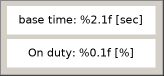
VISUALIZATION vis_FB_DutyCycle_Master  // 164x76
VAR_IN_OUT
	fBaseTime	: REAL;
	fOn_Duty	: REAL;		
END_VAR
    Rectangle (0,0 164x76)
    Textfield (6,5 150x30), "base time: %2.1f [sec]", text variable: fBaseTime
        OnMouseClick: write the text variable via Edit, min 0, max 60
    Textfield (6,38 150x30), "On duty: %0.1f [%]", text variable: fOn_Duty
        OnMouseClick: write the text variable via Edit, min 0, max 100
END_VISUALIZATION

// ---- 01 Instance/04 Recipe/Vis_Recipe_Tab.TcVIS
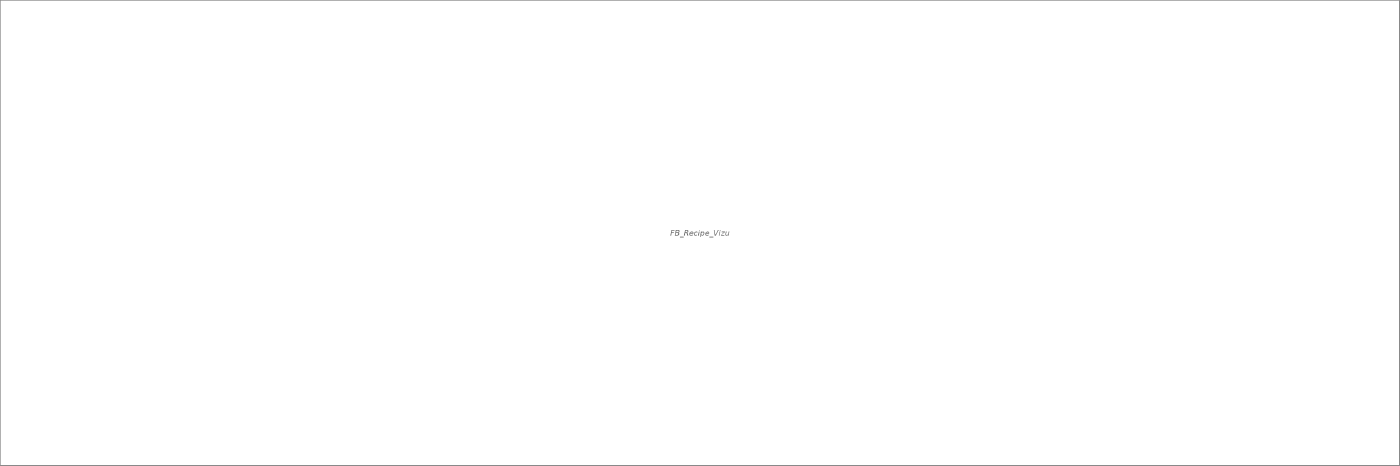
VISUALIZATION Vis_Recipe_Tab  // 1850x617
    TabControl (0,0 1850x617), frame switch variable: prg_Call_Recipe_Slow.iRecipeSwitchFrameVar
        shows FB_Recipe_Vizu(fb_Recipe := GVL_Recipe.fbRecipe[E_Recipe_Name.R_All])
        shows FB_Recipe_Vizu(fb_Recipe := GVL_Recipe.fbRecipe[E_Recipe_Name.R_Device_Dough1])
        shows FB_Recipe_Vizu(fb_Recipe := GVL_Recipe.fbRecipe[E_Recipe_Name.R_Device_Dough2])
        shows FB_Recipe_Vizu(fb_Recipe := GVL_Recipe.fbRecipe[E_Recipe_Name.R_Device_Dough3])
        shows FB_Recipe_Vizu(fb_Recipe := GVL_Recipe.fbRecipe[E_Recipe_Name.R_Device_Dough4])
        shows FB_Recipe_Vizu(fb_Recipe := GVL_Recipe.fbRecipe[E_Recipe_Name.R_CheesyBites])
        shows FB_Recipe_Vizu(fb_Recipe := GVL_Recipe.fbRecipe[E_Recipe_Name.R_CheesyCut])
        shows FB_Recipe_Vizu(fb_Recipe := GVL_Recipe.fbRecipe[E_Recipe_Name.R_Cream])
        shows FB_Recipe_Vizu(fb_Recipe := GVL_Recipe.fbRecipe[E_Recipe_Name.R_Crown])
        shows FB_Recipe_Vizu(fb_Recipe := GVL_Recipe.fbRecipe[E_Recipe_Name.R_Flour])
        shows FB_Recipe_Vizu(fb_Recipe := GVL_Recipe.fbRecipe[E_Recipe_Name.R_Mozzarella])
        shows FB_Recipe_Vizu(fb_Recipe := GVL_Recipe.fbRecipe[E_Recipe_Name.R_Open1])
        shows FB_Recipe_Vizu(fb_Recipe := GVL_Recipe.fbRecipe[E_Recipe_Name.R_Open2])
        shows FB_Recipe_Vizu(fb_Recipe := GVL_Recipe.fbRecipe[E_Recipe_Name.R_Open3])
        shows FB_Recipe_Vizu(fb_Recipe := GVL_Recipe.fbRecipe[E_Recipe_Name.R_Open4])
        shows FB_Recipe_Vizu(fb_Recipe := GVL_Recipe.fbRecipe[E_Recipe_Name.R_Wet])
        shows FB_Recipe_Vizu(fb_Recipe := GVL_Recipe.fbRecipe[E_Recipe_Name.R_Wrap])
        shows FB_Recipe_Vizu(fb_Recipe := GVL_Recipe.fbRecipe[E_Recipe_Name.R_Sesame])
        shows FB_Recipe_Vizu(fb_Recipe := GVL_Recipe.fbRecipe[E_Recipe_Name.R_Piston_Settings])
        [0]: TabTitle=All
        [1]: TabTitle=Device 1
        [2]: TabTitle=Device 2
        [3]: TabTitle=Device 3
        [4]: TabTitle=Device 4
        [5]: TabTitle=Cheesy Bites
        [6]: TabTitle=Cheesy Cut
        [7]: TabTitle=Cream
        [8]: TabTitle=Crown
        [9]: TabTitle=Flour
        [10]: TabTitle=Mozza
        [11]: TabTitle=Open1
        [12]: TabTitle=Open2
        [13]: TabTitle=Open3
        [14]: TabTitle=Open4
        [15]: TabTitle=Wet
        [16]: TabTitle=Wrap
        [17]: TabTitle=Sesame
        [18]: TabTitle=Piston Param
END_VISUALIZATION

// ---- 01 Instance/04-Messages/ERROR_BUFFER.TcVIS
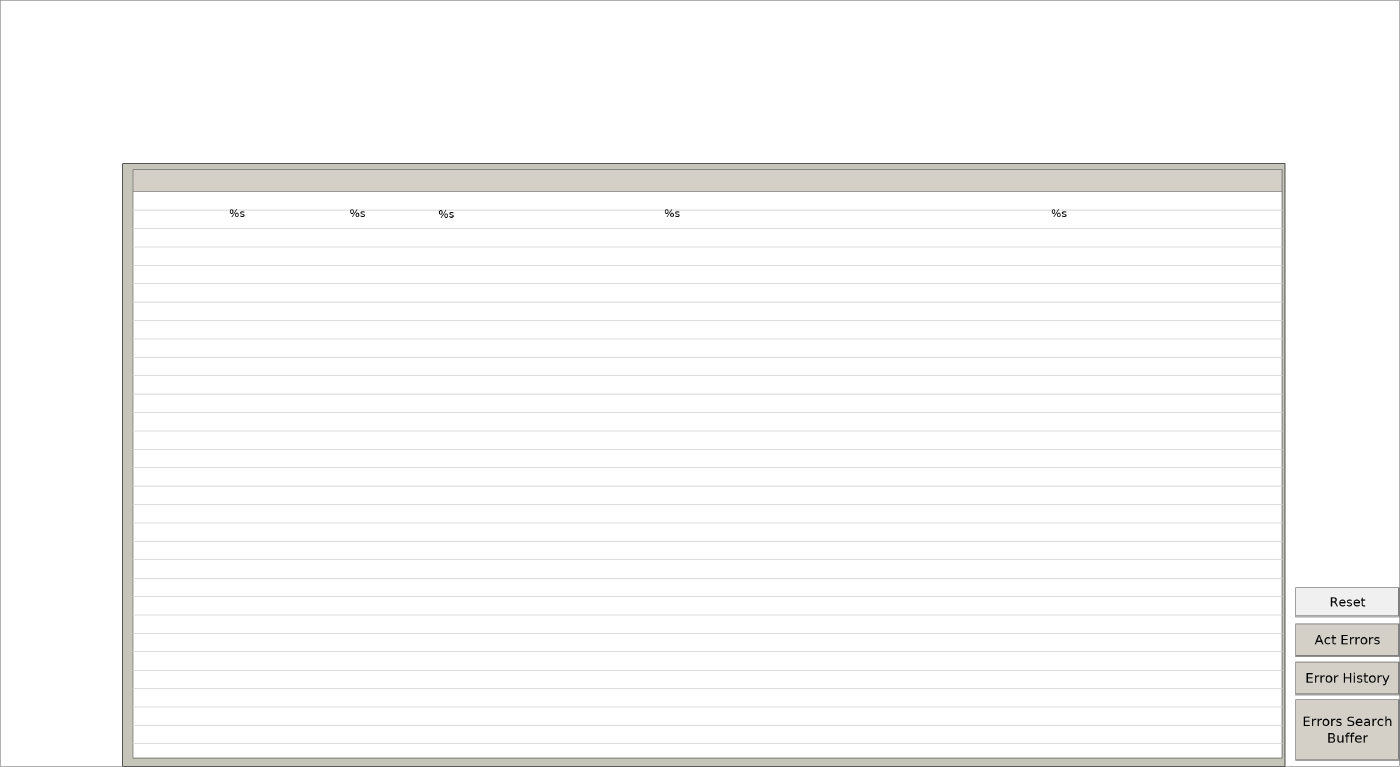
VISUALIZATION ERROR_BUFFER  // 1900x1042
    Group (1758,798 142x235)
        Button (0,0 142x40), "Reset", pressed state: prg_Messages.ResetErrors
            toggle prg_Messages.ResetErrors
        Button (0,101 142x45), "Error History"
            OnMouseClick: change screen: ERROR_HISTORY
        Button (0,152 142x83), "Errors Search Buffer"
            OnMouseClick: change screen: ERROR_BUFFER
        Button (0,49 142x45), "Act Errors"
            OnMouseClick: change screen: ERRORS_OPER
    Rectangle (166,222 1578x820)
    Table (180,230 1560x800), data array: Buffer_Search_Messages
        p3854506369: Buffer_Search_Messages[INDEX].sDateTime
        p1892666644: Buffer_Search_Messages[INDEX].sErrID
        p338671338: Buffer_Search_Messages[INDEX].sLevel
        p2170511999: Buffer_Search_Messages[INDEX].sModuleDescription
        p3723444502: Buffer_Search_Messages[INDEX].sErrorMessage
        p4092479075: Module Description
        p2237128397: Error Message
    Rectangle (421,270 129x40), "%s", text variable: Prg_Filter_Messages.stFilter.sErrID
        OnMouseClick: write the text variable via Edit
    Rectangle (551,271 110x40), "%s", text variable: Prg_Filter_Messages.stFilter.sLevel
        OnMouseClick: write the text variable via Edit
    Rectangle (662,270 501x40), "%s", text variable: Prg_Filter_Messages.stFilter.sModuleDescription
        OnMouseClick: write the text variable via Edit
    Rectangle (1162,270 551x40), "%s", text variable: Prg_Filter_Messages.stFilter.sErrorMessage
        OnMouseClick: write the text variable via Edit
    Rectangle (222,270 200x40), "%s", text variable: Prg_Filter_Messages.stFilter.sDateTime
        OnMouseClick: write the text variable via Edit
END_VISUALIZATION

// ---- 01 Instance/04-Messages/ERROR_HISTORY.TcVIS
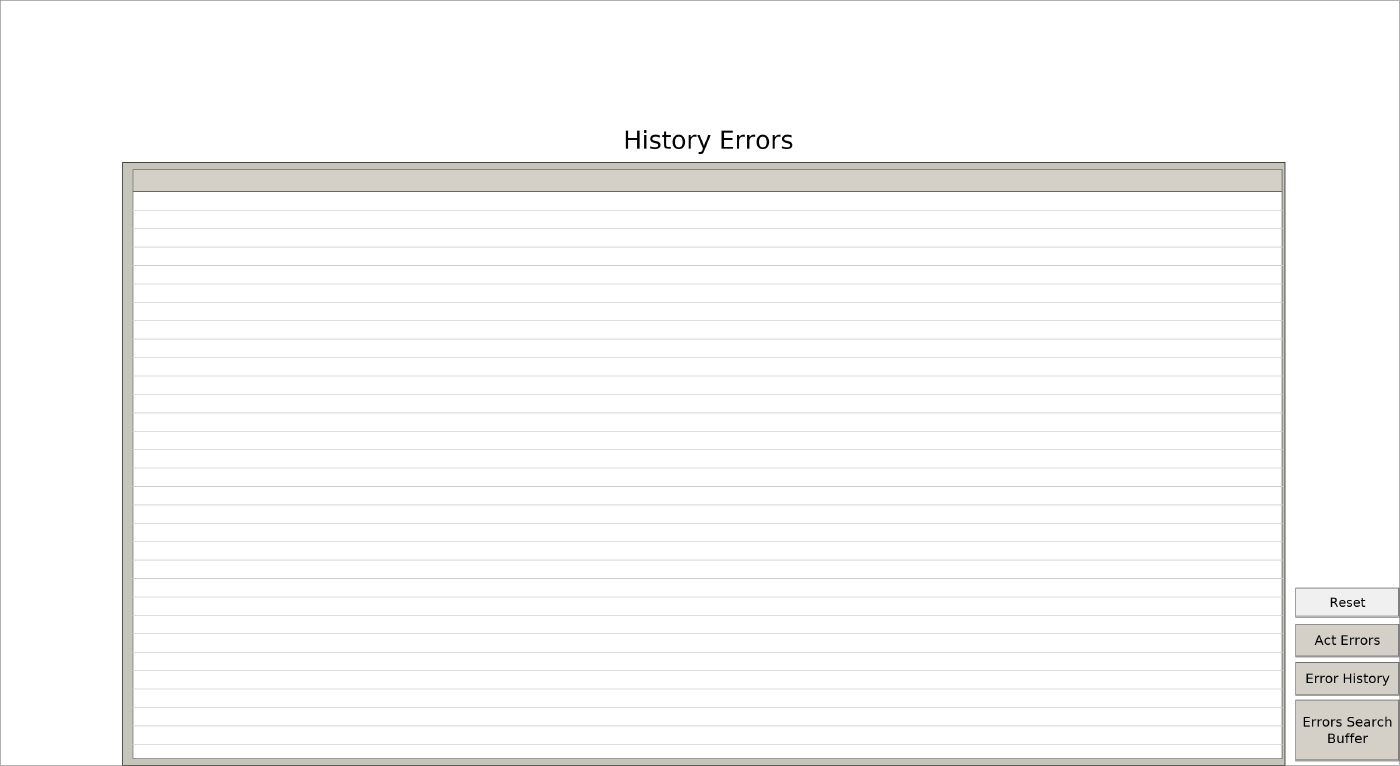
VISUALIZATION ERROR_HISTORY  // 1900x1040
    Group (1758,798 142x235)
        Button (0,0 142x40), "Reset", pressed state: prg_Messages.ResetErrors
            toggle prg_Messages.ResetErrors
        Button (0,101 142x45), "Error History"
            OnMouseClick: change screen: ERROR_HISTORY
        Button (0,152 142x83), "Errors Search Buffer"
            OnMouseClick: change screen: ERROR_BUFFER
        Button (0,49 142x45), "Act Errors"
            OnMouseClick: change screen: ERRORS_OPER
    Rectangle (166,220 1578x820)
    Rectangle (841,165 241x50), "History Errors"
    Table (180,230 1560x800), data array: Buffer_Act_History
        p3854506369: Buffer_Act_History[INDEX].sDateTime
        p1892666644: Buffer_Act_History[INDEX].sErrID
        p338671338: Buffer_Act_History[INDEX].sLevel
        p2170511999: Buffer_Act_History[INDEX].sModuleDescription
        p3723444502: Buffer_Act_History[INDEX].sErrorMessage
        p4092479075: Module Description
        p2237128397: Error Message
END_VISUALIZATION

// ---- 01 Instance/04-Messages/ERROR_Tab.TcVIS
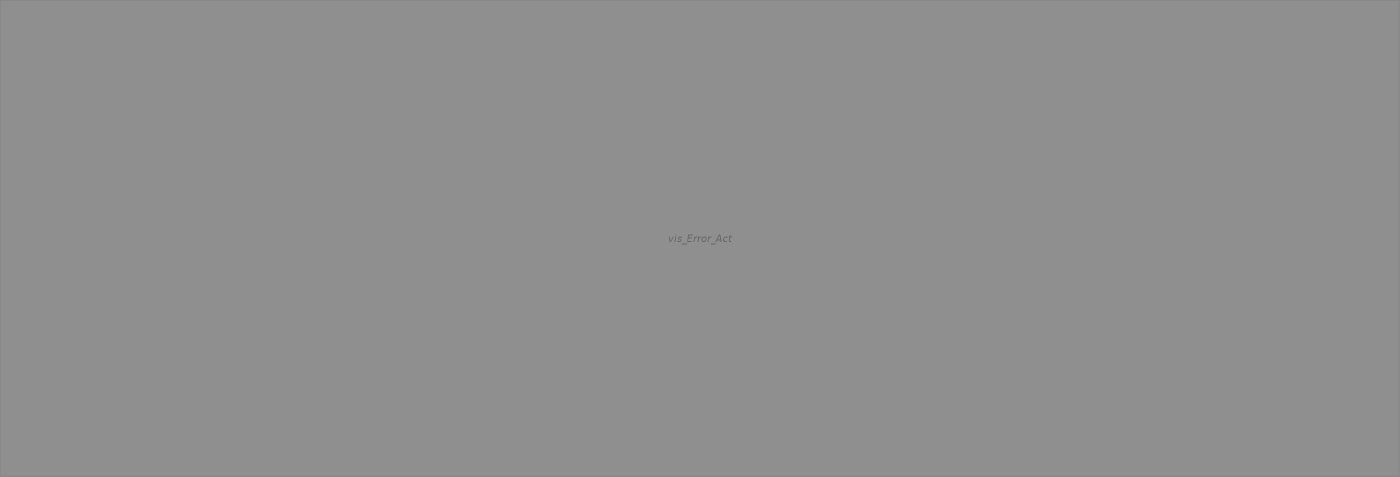
VISUALIZATION ERROR_Tab  // 1428x487
    Rectangle (0,0 1428x487)
    TabControl (0,0 1428x487)
        shows vis_Error_Act()
        shows vis_Error_History()
        shows vis_Error_Search()
        [0]: TabTitle=Actual Errors
        [1]: TabTitle=Error History
        [2]: TabTitle=Search
END_VISUALIZATION

// ---- 01 Instance/04-Messages/ERROR_Tab_1.TcVIS
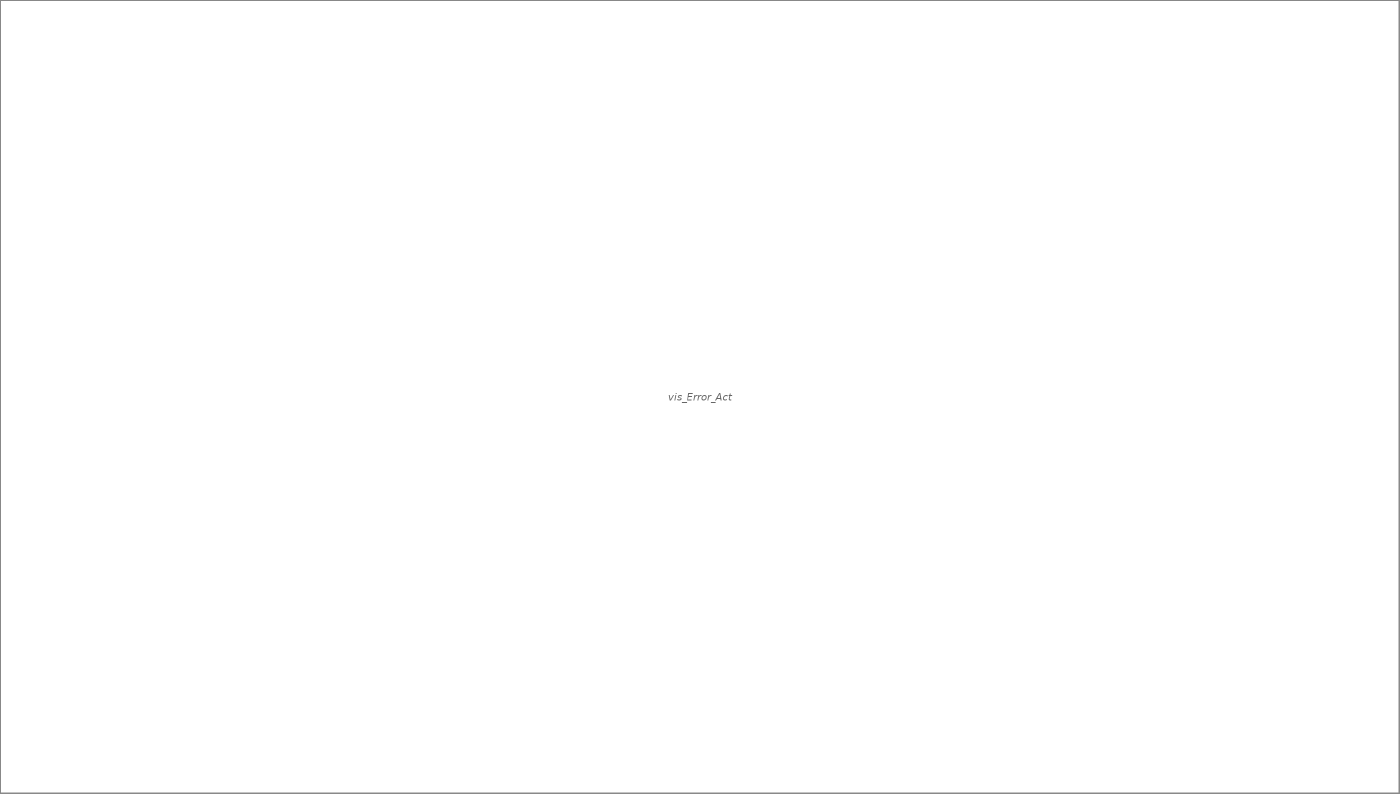
VISUALIZATION ERROR_Tab_1  // 1428x810
    TabControl (0,0 1428x810)
        shows vis_Error_Act()
        shows vis_Error_History()
        shows vis_Error_Search()
        [0]: TabTitle=Actual
        [1]: TabTitle=History
        [2]: TabTitle=Search
END_VISUALIZATION

// ---- 01 Instance/04-Messages/vis_Error_Act.TcVIS
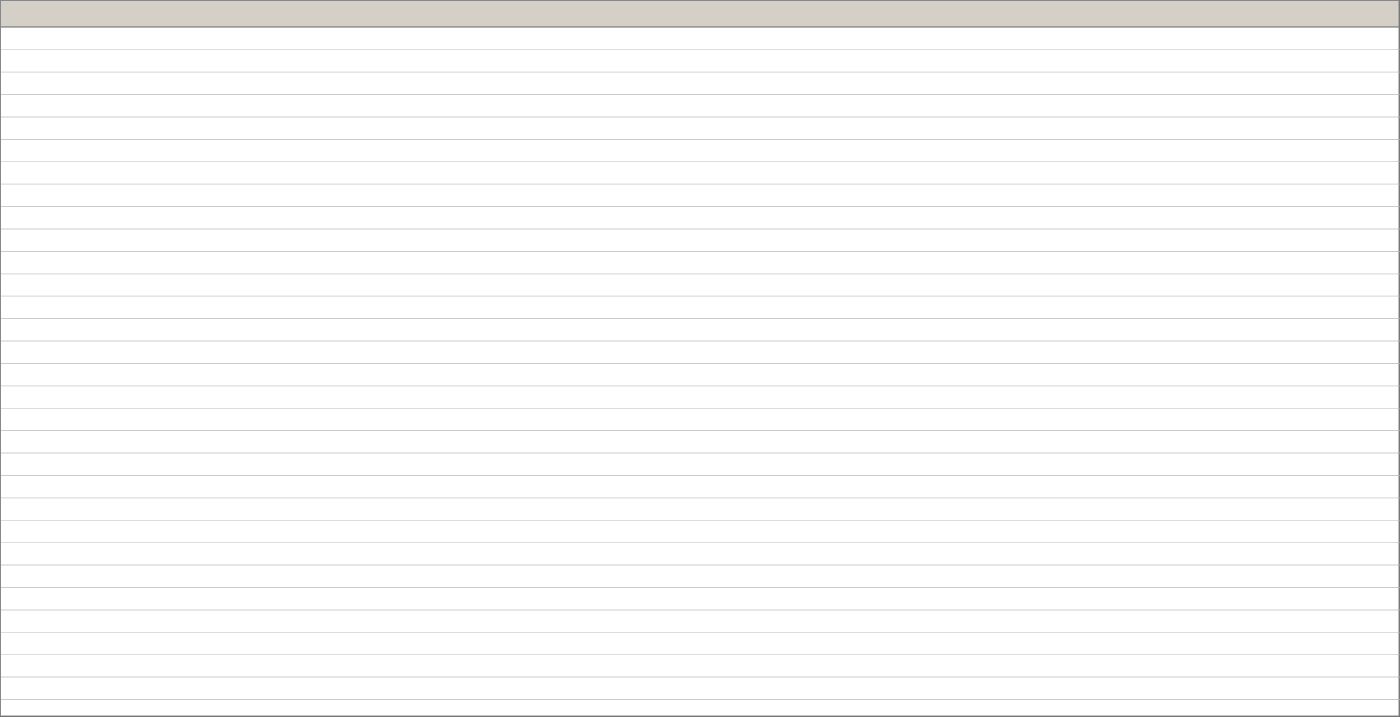
VISUALIZATION vis_Error_Act  // 1560x800
    Table (0,0 1560x800), data array: Buffer_Act_Message
        p3854506369: Buffer_Act_Message[INDEX].sDateTime
        p1892666644: Buffer_Act_Message[INDEX].sErrID
        p338671338: Buffer_Act_Message[INDEX].sLevel
        p2170511999: Buffer_Act_Message[INDEX].sModuleDescription
        p3723444502: Buffer_Act_Message[INDEX].sErrorMessage
        p4092479075: Module Description
        p2237128397: Error Message
END_VISUALIZATION

// ---- 01 Instance/04-Messages/vis_Error_History.TcVIS
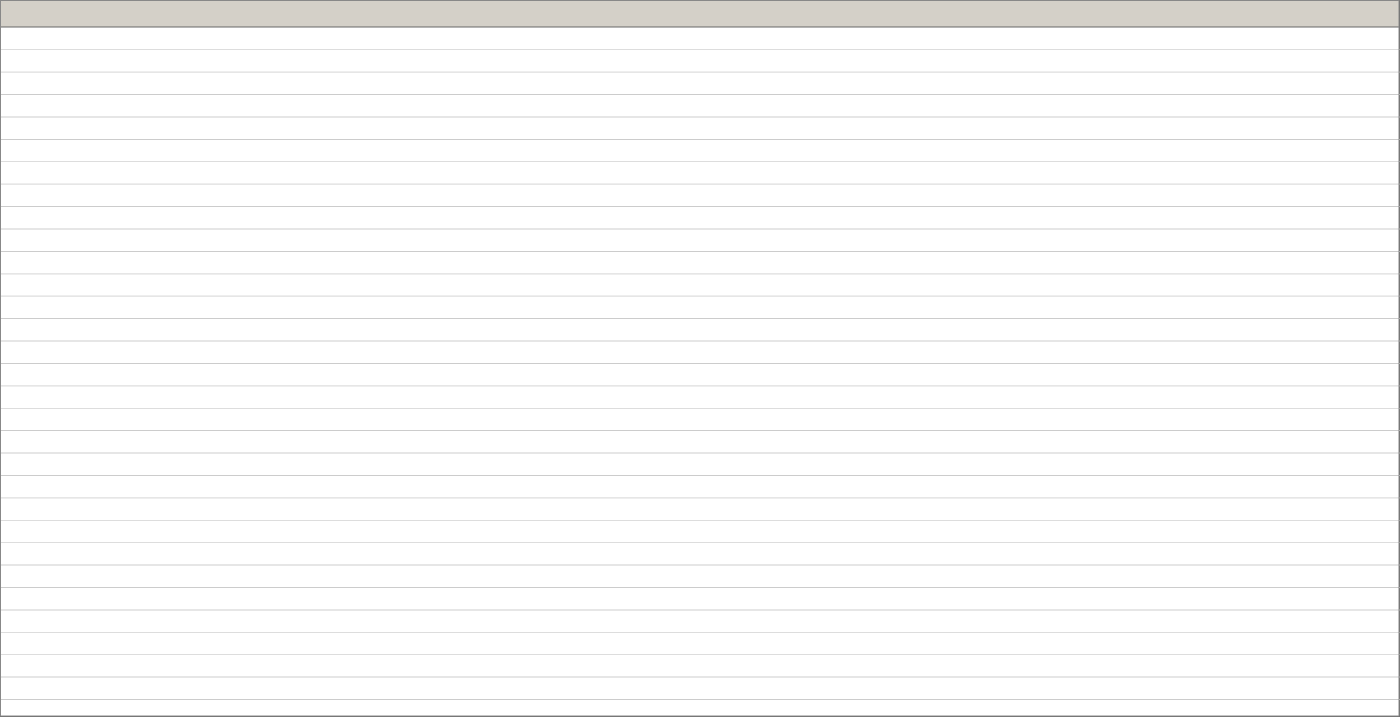
VISUALIZATION vis_Error_History  // 1560x800
    Table (0,0 1560x800), data array: Buffer_Act_History
        p3854506369: Buffer_Act_History[INDEX].sDateTime
        p1892666644: Buffer_Act_History[INDEX].sErrID
        p338671338: Buffer_Act_History[INDEX].sLevel
        p2170511999: Buffer_Act_History[INDEX].sModuleDescription
        p3723444502: Buffer_Act_History[INDEX].sErrorMessage
        p4092479075: Module Description
        p2237128397: Error Message
END_VISUALIZATION

// ---- 01 Instance/04-Messages/vis_Error_Search.TcVIS
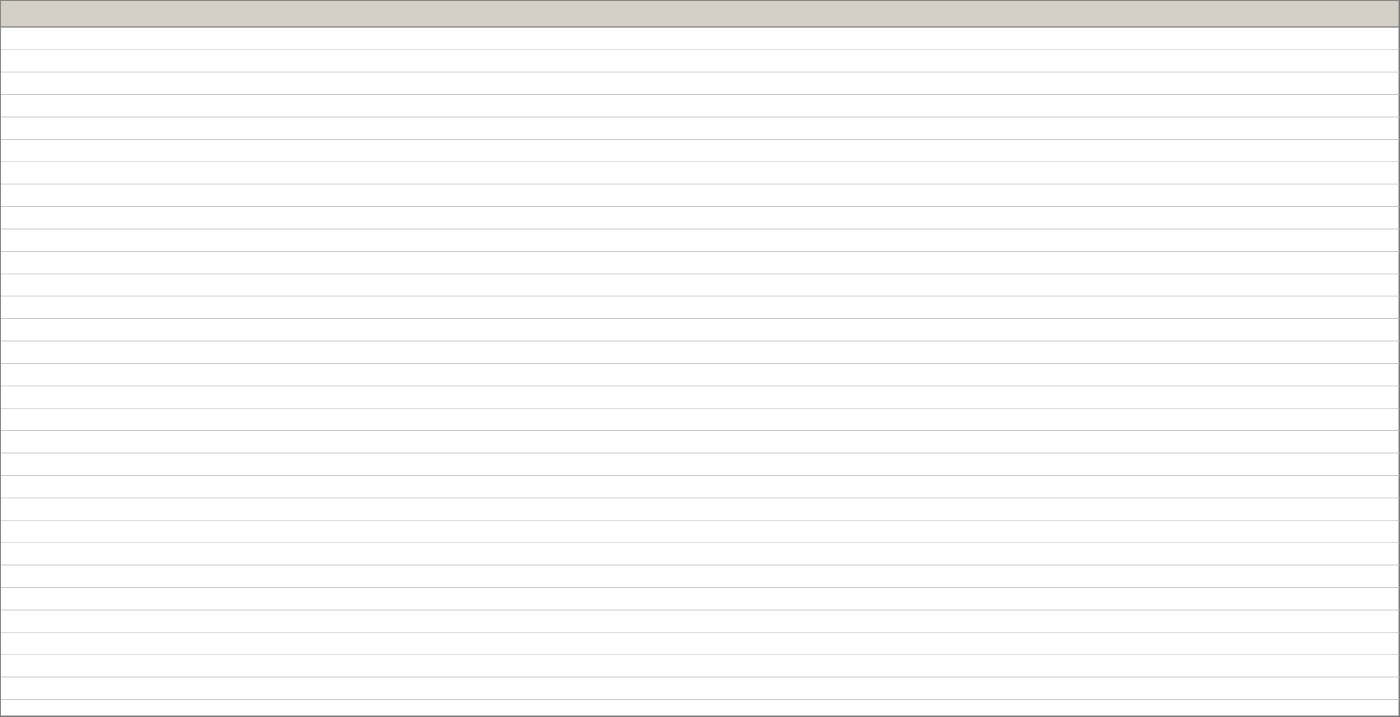
VISUALIZATION vis_Error_Search  // 1560x800
    Table (0,0 1560x800), data array: Buffer_Search_Messages
        p3854506369: Buffer_Search_Messages[INDEX].sDateTime
        p1892666644: Buffer_Search_Messages[INDEX].sErrID
        p338671338: Buffer_Search_Messages[INDEX].sLevel
        p2170511999: Buffer_Search_Messages[INDEX].sModuleDescription
        p3723444502: Buffer_Search_Messages[INDEX].sErrorMessage
        p4092479075: Module Description
        p2237128397: Error Message
END_VISUALIZATION

// ---- 01 Instance/06-Visu/ERRORS_OPER_16_9.TcVIS
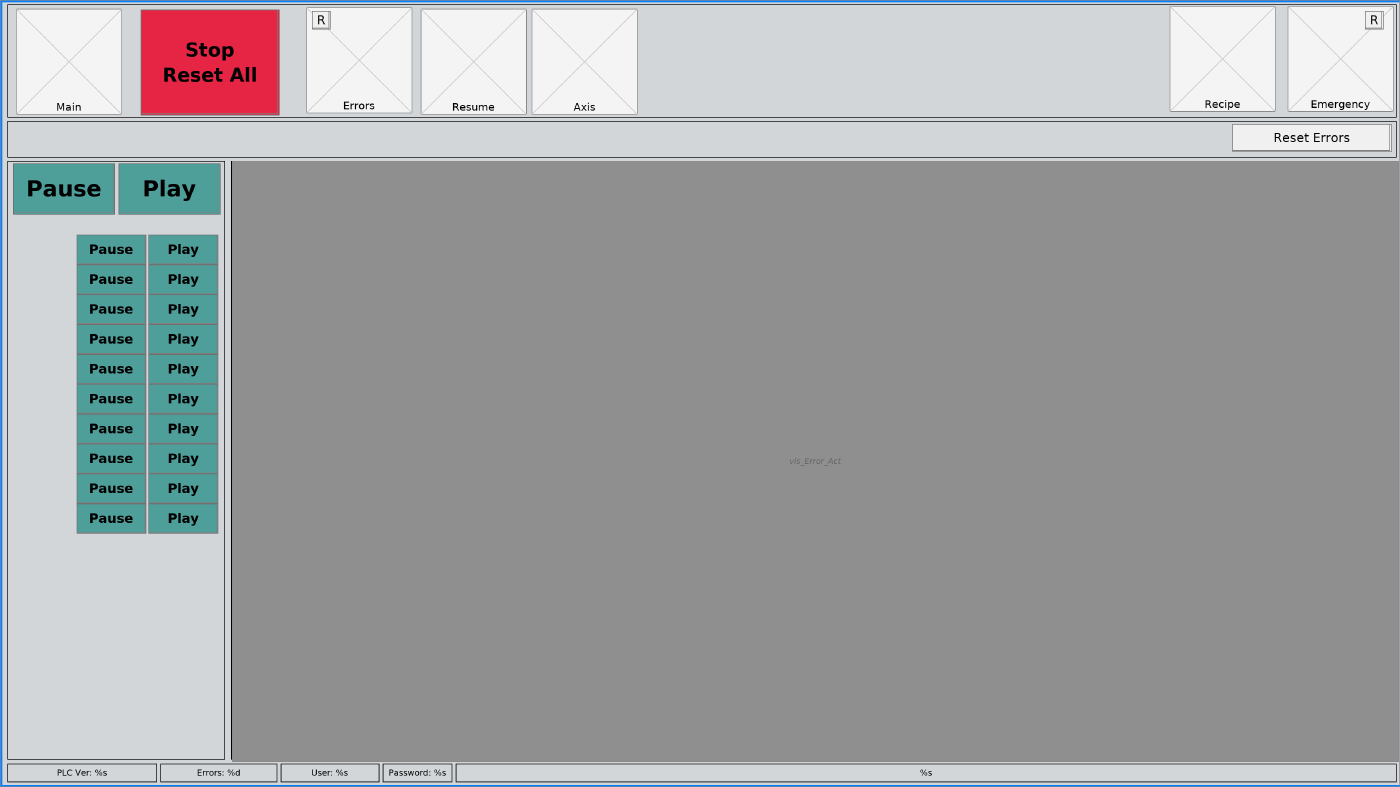
VISUALIZATION ERRORS_OPER_16_9  // 1920x1080
    Frame (0,0 1920x1080)
        shows TEMP16_9_00()
    Frame (318,221 1600x824)
        shows ERROR_Tab()
    Button (1690,170 218x38), "Reset Errors", pressed state: prg_Messages.ResetErrors
        toggle prg_Messages.ResetErrors
END_VISUALIZATION

// ---- 01 Instance/06-Visu/ES_INT_OPER_16_9.TcVIS
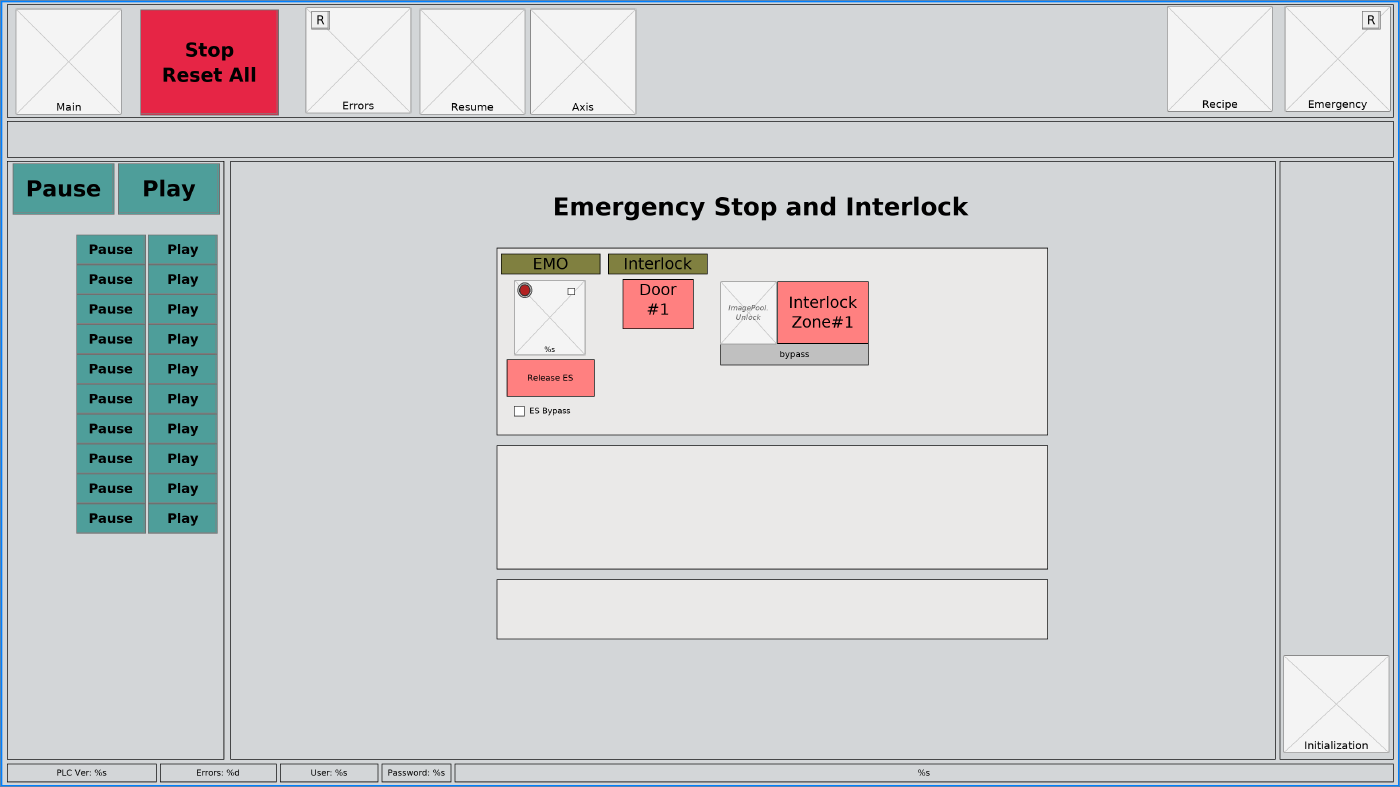
VISUALIZATION ES_INT_OPER_16_9  // 1920x1080
    Frame (0,0 1920x1080)
        shows TEMP16_9_00()
    Rectangle (742,266 602x35), "Emergency Stop and Interlock"
    Rectangle (681,611 756x170)
    Rectangle (681,340 756x257)
    Rectangle (681,795 756x82), invisible if: prg_User.actUser<4
    Rectangle (695,493 120x51), "Release ES", colour toggle: bStateSafe
    Checkbox (703,552 111x24), "ES Bypass", variable: bES_Bypass, invisible if: prg_User.actUser<4
    RoundedRectangle (687,348 136x28), "EMO"
    Frame (705,384 100x103)
        shows Vis_ES_PB(stPB := bES_PB[1], Lable := 'EMO#1')
    RoundedRectangle (834,348 136x28), "Interlock"
    Rectangle (854,383 97x68), "Door #1", colour toggle: bInterlock[1]
    Group (988,386 203x115)
        Rectangle (78,0 125x85), "Interlock Zone#1", colour toggle: bIntZoneLocked[1]
        Rectangle (0,85 203x30), "bypass", colour toggle: bIntZoneBypass[1], invisible if: NOT bIntZoneBypass[1]
            toggle bIntZoneBypass[1]
        Image (0,0 77x86), input disabled if: prg_User.actUser<3, image: ImagePool.Unlock
            p84334746: GVL_Safety.sInterlocksZone1
            OnMouseClick: toggle bIntZoneBypass[1]
END_VISUALIZATION

// ---- 01 Instance/06-Visu/Recipe_16_9.TcVIS
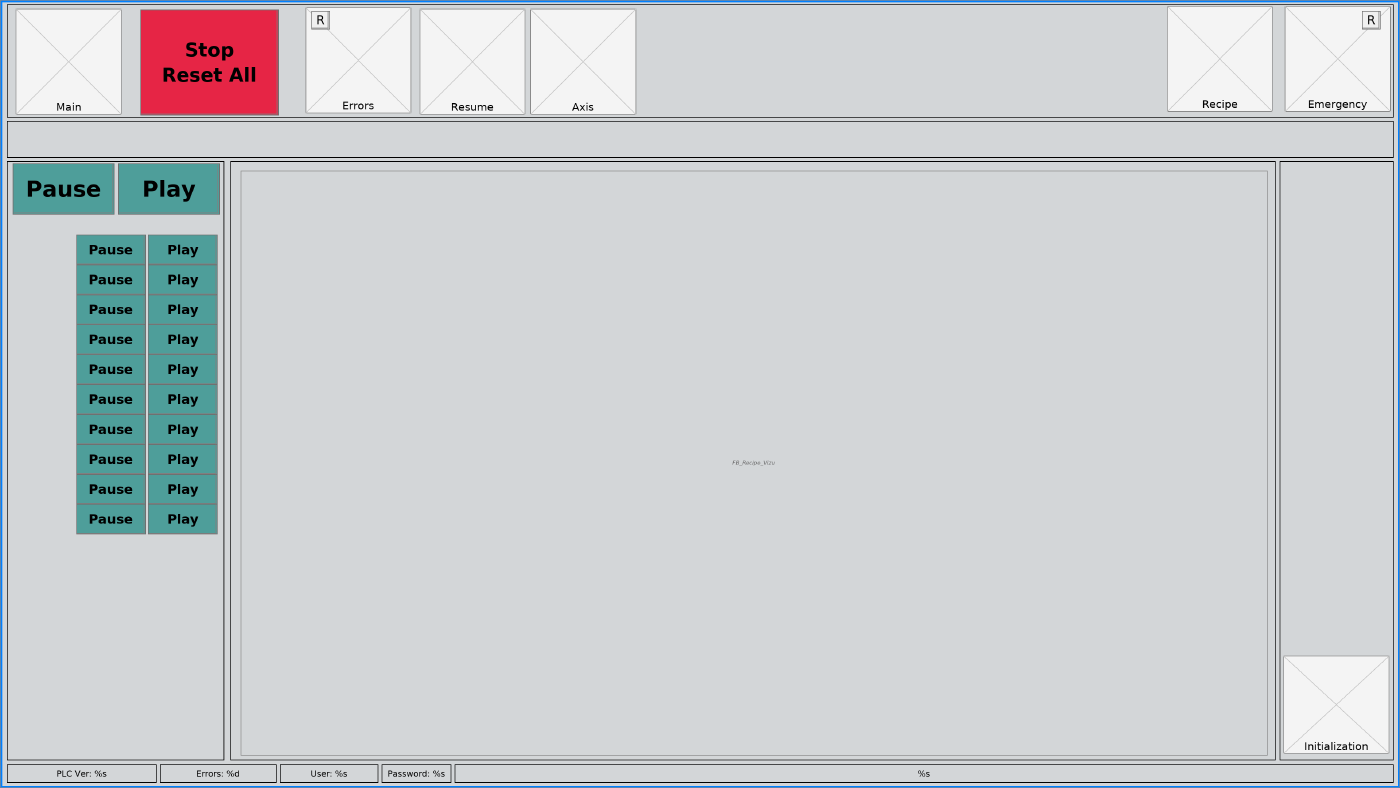
VISUALIZATION Recipe_16_9  // 1920x1081
    Frame (0,0 1920x1081)
        shows TEMP16_9_00()
    Frame (330,234 1408x802)
        shows Vis_Recipe_Tab()
END_VISUALIZATION

// ---- 01 Instance/06-Visu/Template16-9/TEMP16_9_00.TcVIS
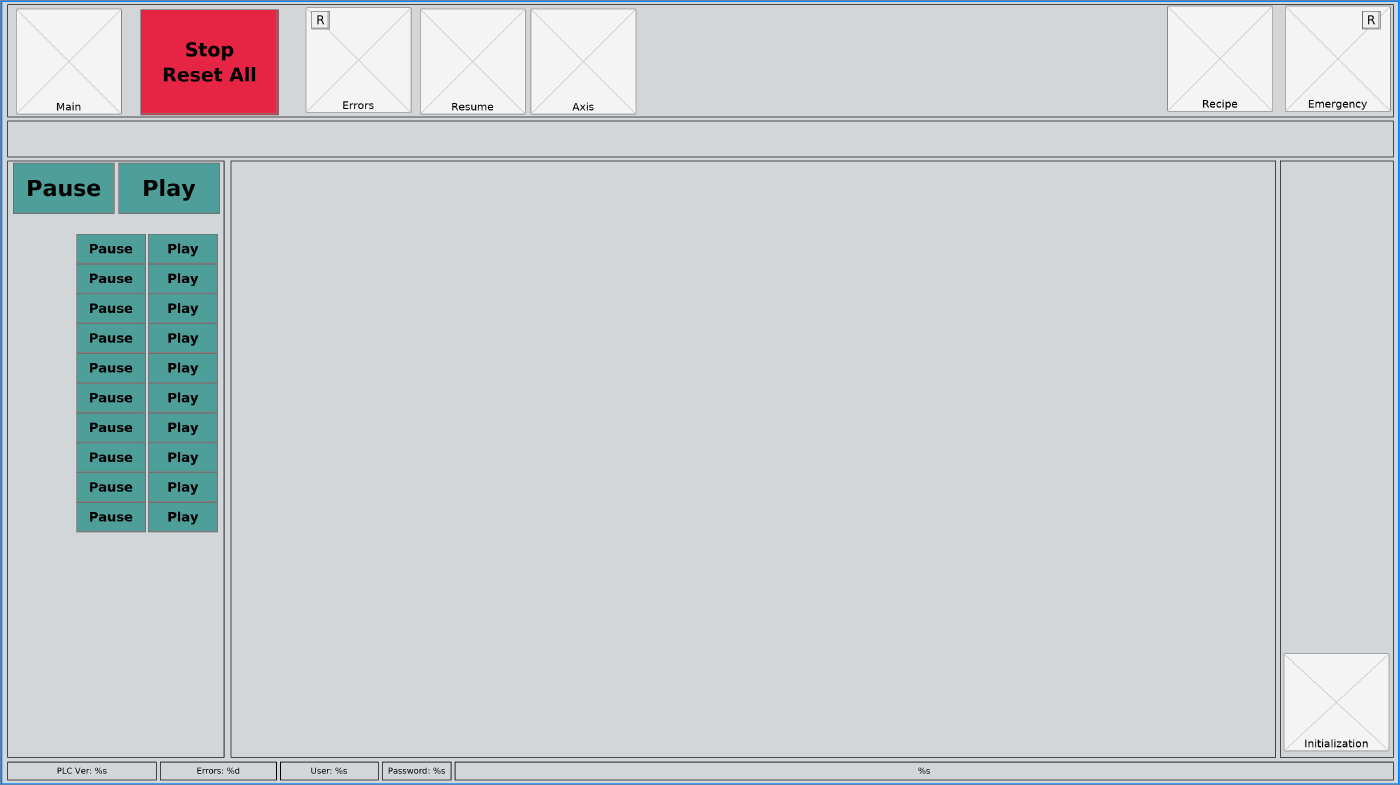
VISUALIZATION TEMP16_9_00  // 1924x1080
    Rectangle (0,0 1924x1080)
    Rectangle (385,1048 135x25), "User: %s", text variable: prg_User.actUser
    Rectangle (525,1048 95x25), "Password: %s", text variable: prg_User.Password
        OnMouseDown: write the text variable via Edit, min 1, max 999
    Rectangle (220,1048 160x25), "Errors: %d", text variable: Global_Persistent.Errors, colour toggle: Global_Persistent.Errors<>0
        OnMouseUp: execute { Global_Persistent.Errors:=(0); }
    Rectangle (10,1048 205x25), "PLC Ver: %s", text variable: ProgramVersion
    Rectangle (625,1048 1290x25), "%s", text variable: sDateTime
    Rectangle (10,6 1905x155)
    Rectangle (10,166 1905x50)
    Image (22,12 145x145), "Main", image: ImagePool.Main
        OnMouseClick: change screen: vis_MAIN
    Image (1766,8 145x145), "Emergency", image: ImagePool.EStop_OK2
        p84334746: GVL_Safety.sBitmap_ESButton
        OnMouseClick: change screen: ES_INT_OPER_16_9
    Image (420,10 145x145), "Errors", image: ImagePool.Error_No
        p84334746: s_Error_BitmapID
        OnMouseClick: change screen: ERRORS_OPER_16_9
    Image (577,12 145x145), "Resume", image: ImagePool.Resume3
        OnMouseClick: toggle ResumeAll
    Button (428,15 25x25), "R", pressed state: prg_Messages.ResetErrors
        toggle prg_Messages.ResetErrors
    Button (1872,15 25x25), "R"
    Rectangle (10,221 298x821)
    Rectangle (1759,221 156x821)
    Frame (18,224 284x70)
        shows OperationButtons(stOperation := stOpMain)
    Image (1764,899 145x134), "Initialization", image: ImagePool.illustration-project-icon
        OnMouseClick: change screen: INIT_OPER_16_9
    Rectangle (317,221 1436x821)
    Frame (193,13 190x145)
        shows OperationButton_Stop(stOperation := stOpMain)
    Image (729,12 145x145), "Axis", image: ImagePool.ervo-motor-beckhoff
        OnMouseClick: change screen: AXIS_OPER
    Image (1604,8 145x145), "Recipe", image: ImagePool.recipe icon
        OnMouseClick: change screen: Recipe_16_9
    Frame (105,322 194x41)
        shows OperationButtons(stOperation := stOper[E_ModeZone.eMain])
    Frame (105,363 194x41)
        shows OperationButtons(stOperation := stOper[E_ModeZone.eCIP])
    Frame (105,404 194x41)
        shows OperationButtons(stOperation := stOper[E_ModeZone.eTank1])
    Frame (105,445 194x41)
        shows OperationButtons(stOperation := stOper[E_ModeZone.eTank2])
    Frame (105,486 194x41)
        shows OperationButtons(stOperation := stOper[E_ModeZone.eTank3])
    Frame (105,527 194x41)
        shows OperationButtons(stOperation := stOper[E_ModeZone.eTank4])
    Frame (105,568 194x41)
        shows OperationButtons(stOperation := stOper[E_ModeZone.eProduction_Marinade])
    Frame (105,609 194x41)
        shows OperationButtons(stOperation := stOper[E_ModeZone.eProduction_Color])
    Frame (105,650 194x41)
        shows OperationButtons(stOperation := stOper[E_ModeZone.eTriBlender_Marinade])
    Frame (105,691 194x41)
        shows OperationButtons(stOperation := stOper[E_ModeZone.eTriBlender_Color])
END_VISUALIZATION

// ---- 01 Instance/06-Visu/Template16-9/TEMP16_9_00_1.TcVIS
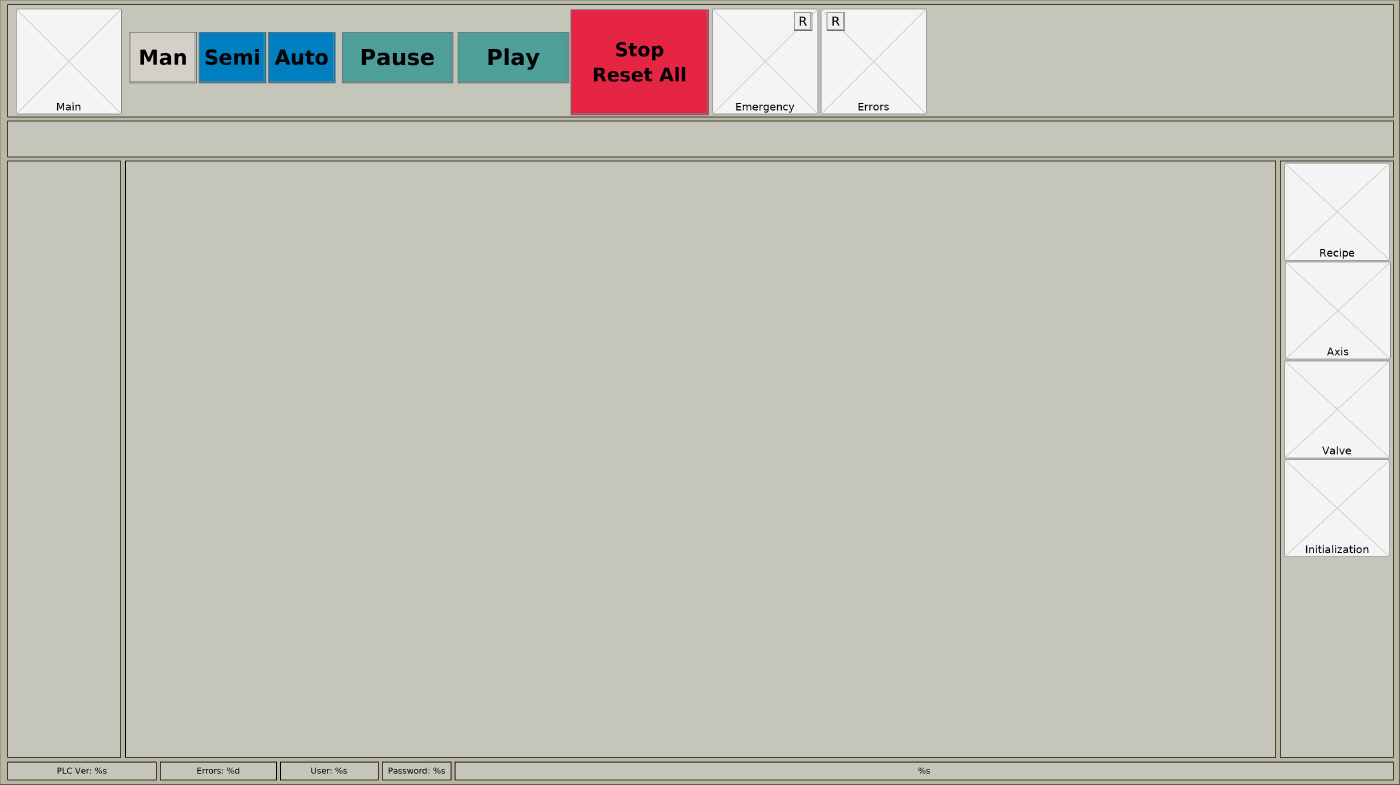
VISUALIZATION TEMP16_9_00_1  // 1924x1080
    Rectangle (0,0 1924x1080)
    Rectangle (385,1048 135x25), "User: %s", text variable: prg_User.actUser
    Rectangle (525,1048 95x25), "Password: %s", text variable: prg_User.Password
        OnMouseDown: write the text variable via Default, min 1, max 999
    Rectangle (220,1048 160x25), "Errors: %d", text variable: Global_Persistent.Errors, colour toggle: Global_Persistent.Errors<>0
        OnMouseUp: execute { Global_Persistent.Errors:=(0); }
    Rectangle (10,1048 205x25), "PLC Ver: %s", text variable: ProgramVersion
    Rectangle (625,1048 1290x25), "%s", text variable: sDateTime
    Rectangle (10,6 1905x155)
    Rectangle (10,166 1905x50)
    Image (22,12 145x145), "Main", image: ImagePool.Main
        OnMouseClick: change screen: vis_MAIN
    Image (979,12 145x145), "Emergency", image: ImagePool.EStop_OK2
        p84334746: GVL_Safety.sBitmap_ESButton
        OnMouseClick: change screen: ES_INT_OPER_16_9
    Image (1128,12 145x145), "Errors", image: ImagePool.Error_No
        p84334746: s_Error_BitmapID
        OnMouseClick: change screen: ERRORS_OPER_16_9
    Button (1136,17 25x25), "R", pressed state: prg_Messages.ResetErrors
        toggle prg_Messages.ResetErrors
    Button (1091,17 25x25), "R"
    Rectangle (10,221 156x821)
    Rectangle (1759,221 156x821)
    Image (1765,224 145x134), "Recipe", image: ImagePool.recipe icon
        OnMouseClick: change screen: Recipe_16_9
    Image (1765,496 145x134), "Valve", image: ImagePool.festo-pistonjpg
        OnMouseClick: change screen: PISTON_OPER_16_9
    Frame (470,44 312x70)
        shows OperationButtons(stOperation := stOpMain)
    Frame (178,44 283x70)
        shows Mode_Select(stMode := stModeMain)
    Image (1765,632 145x134), "Initialization", image: ImagePool.illustration-project-icon
        OnMouseClick: change screen: INIT_OPER_16_9
    Rectangle (172,221 1581x821)
    Frame (784,13 190x145)
        shows OperationButton_Stop(stOperation := stOpMain)
    Image (1766,360 145x134), "Axis", image: ImagePool.ervo-motor-beckhoff
        OnMouseClick: change screen: AXIS_OPER
END_VISUALIZATION

// ---- 01 Instance/06-Visu/Template16-9/TEMP16_9_00_Content.TcVIS
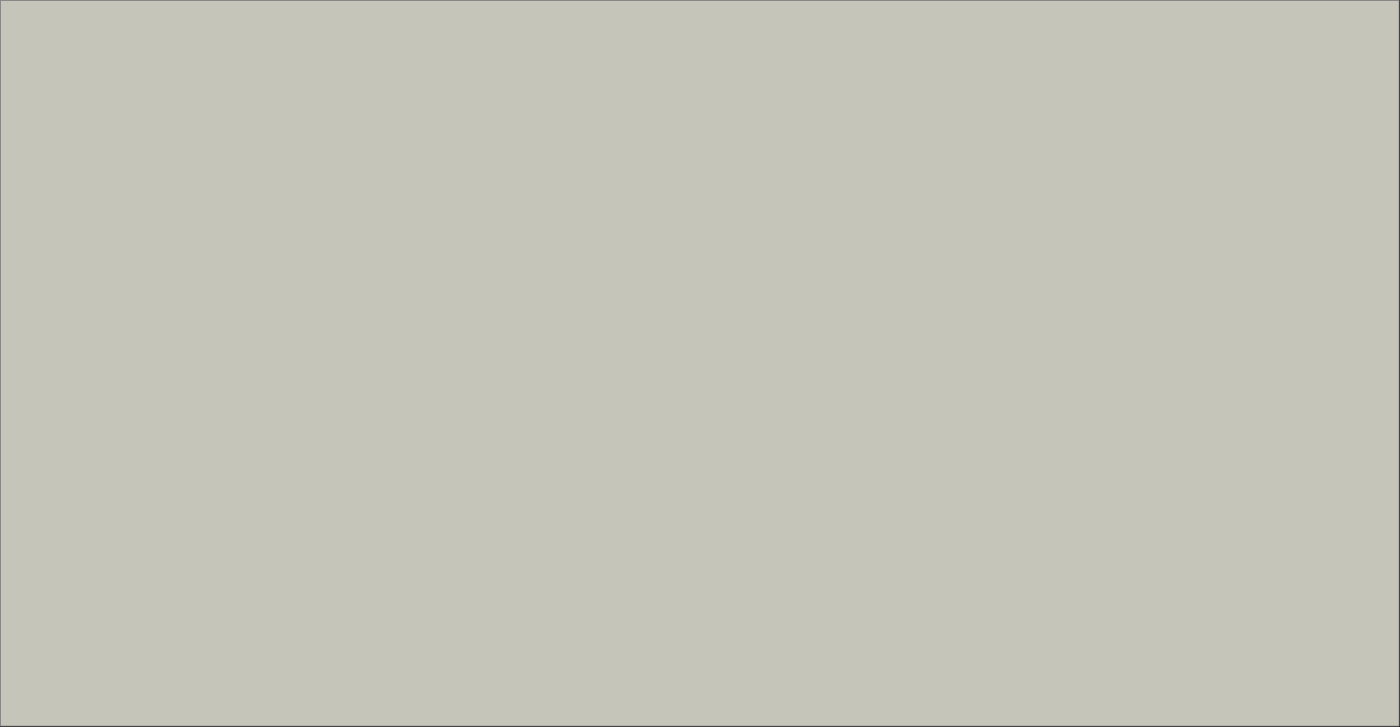
VISUALIZATION TEMP16_9_00_Content  // 1581x821
    Rectangle (0,0 1581x821)
END_VISUALIZATION

// ---- 01 Instance/07-Mode/Vis_LightTower.TcVIS
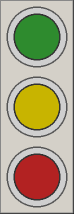
VISUALIZATION Vis_LightTower  // 74x214
    Rectangle (0,0 74x214), colour toggle: prg_LightTower.qBuzzer
    Lamp1 (2,2 70x70), variable: prg_LightTower.qLedGreen, style: Lamp-Lamp1-Green
    Lamp1 (2,72 70x70), variable: prg_LightTower.qLedYellow, style: Lamp-Lamp1-Yellow
    Lamp1 (2,142 70x70), variable: prg_LightTower.qLedRed, style: Lamp-Lamp1-Red
END_VISUALIZATION

// ---- 01 Instance/07-Mode/Vis_LightTower_1.TcVIS
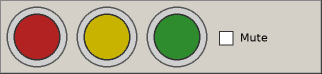
VISUALIZATION Vis_LightTower_1  // 322x74
    Rectangle (0,0 322x74), colour toggle: prg_LightTower.qBuzzer
    Group (2,2 210x70)
        Lamp1 (140,0 70x70), variable: prg_LightTower.qLedGreen, style: Lamp-Lamp1-Green
        Lamp1 (70,0 70x70), variable: prg_LightTower.qLedYellow, style: Lamp-Lamp1-Yellow
        Lamp1 (0,0 70x70), variable: prg_LightTower.qLedRed, style: Lamp-Lamp1-Red
    Checkbox (217,13 95x50), "Mute", variable: bBuzzerMute, input disabled if: prg_User.actUser<2
END_VISUALIZATION

// ---- 01 Instance/07-Mode/viz_HMI_LockIndex.TcVIS
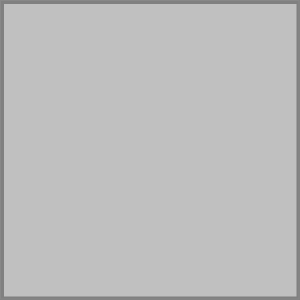
VISUALIZATION viz_HMI_LockIndex  // 300x300
    Rectangle (0,0 300x300), invisible if: not prg_HMI_OperationLock.b_LockIndex
END_VISUALIZATION

// ---- 01 Instance/07-Mode/viz_HMI_Piston.TcVIS
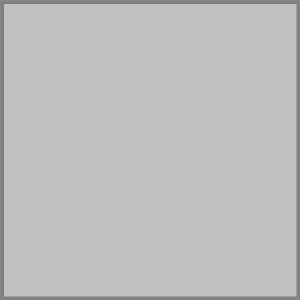
VISUALIZATION viz_HMI_Piston  // 300x300
VAR_INPUT
	bLock_HMI: BOOL;
END_VAR
    Rectangle (0,0 300x300), invisible if: TRUE
END_VISUALIZATION

// ---- 03 Project/10 Element/TextList_InterConnection.TcTLO
TEXTLIST TextList_InterConnection
  0 = 'Not Connected'
  1 = 'TriBlender'
  2 = 'Production Line'
  3 = 'Tank'
  4 = 'CIP'
   = ''
END_TEXTLIST

// ---- 03 Project/10 Element/TextList_StateLong.TcTLO
TEXTLIST TextList_StateLong
  0 = 'Off'
  1 = 'Standby'
  2 = 'Not Clean'
  3 = 'CIP1 - Rinzed'
  4 = 'CIP2 - Deterged'
  5 = 'CIP3 - Deterged + Clean'
  6 = 'CIP4 - Disinfected'
  7 = 'CIP5 - Done'
  8 = 'Water Ready'
  9 = 'Ready'
  10 = 'Production'
  11 = 'Empty'
  12 = 'Expired'
   = ''
END_TEXTLIST

// ---- 03 Project/10 Element/TextList_StateLong_1.TcTLO
TEXTLIST TextList_StateLong_1
  0 = 'Not Clean'
  7 = 'Clean'
  9 = 'Product'
   = ''
END_TEXTLIST

// ---- 03 Project/10 Element/vis_FB_Element.TcVIS
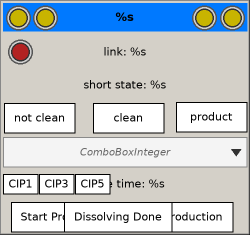
VISUALIZATION vis_FB_Element  // 250x235
VAR_IN_OUT
	fb: FB_Element;
END_VAR
    Rectangle (0,0 250x235)
    Textfield (3,70 244x30), "short state: %s", text variable: fb.eState_Short
    ComboBoxInteger (3,137 244x30), variable: fb.eState_Long, input disabled if: fb.bStateUpdate_Limited, text list: 'TextList_StateLong'
    Textfield (2,2 246x30), "%s", text variable: fb.sElementID
    Textfield (2,169 246x30), "state time: %s", text variable: fb.sState_Time
    RoundedRectangle (11,202 108x30), "Start Production", invisible if: NOT (fb.eInterConnect=E_InterConnection.ConnToLine AND fb.eState_Long=E_Element_State_Long.eReady)
        OnMouseClick: execute { fb.eState_Long:=E_Element_State_Long.eProduction; }
    RoundedRectangle (125,202 108x30), "Stop Production", invisible if: NOT (fb.eInterConnect=E_InterConnection.ConnToLine AND fb.eState_Long=E_Element_State_Long.eProduction)
        OnMouseClick: execute { fb.eState_Long:=E_Element_State_Long.eReady; }
    RoundedRectangle (64,202 108x30), "Dissolving Done", invisible if: NOT ((fb.eInterConnect=E_InterConnection.ConnToTriBlender) AND (fb.eState_Long=E_Element_State_Long.eCIP_5_Done OR fb.eState_Long=E_Element_State_Long.eWaterReady))
        OnMouseClick: execute { fb.eState_Long:=E_Element_State_Long.eReady; }
    Lamp1 (190,4 29x28), variable: fb.eInterConnect=E_InterConnection.ConnToLine, style: Lamp-Lamp1-Yellow
    Lamp1 (218,4 29x28), variable: fb.eInterConnect=E_InterConnection.ConnToTriBlender, style: Lamp-Lamp1-Yellow
    Lamp1 (31,4 29x28), variable: fb.eInterConnect=E_InterConnection.ConnToTank, style: Lamp-Lamp1-Yellow
    Textfield (3,37 244x30), "link: %s", colour toggle: fb.eInterConnect<>0, text list: 'TextList_InterConnection', text index: fb.eInterConnect
    RoundedRectangle (4,103 71x30), "not clean"
        OnMouseClick: execute { fb.eState_Long:=E_Element_State_Long.eNotClean; }
    RoundedRectangle (93,103 71x30), "clean"
        OnMouseClick: execute { fb.eState_Long:=E_Element_State_Long.eCIP_5_Done; }
    RoundedRectangle (176,102 71x30), "product"
        OnMouseClick: execute { fb.eState_Long:=E_Element_State_Long.eProduction; }
    Lamp1 (4,4 29x28), variable: fb.eInterConnect=E_InterConnection.ConnToCIP, style: Lamp-Lamp1-Yellow
    RoundedRectangle (3,174 35x20), "CIP1"
        tap fb.bTakePosInCIPBuffer_Partial
    RoundedRectangle (39,174 35x20), "CIP3"
        tap fb.bTakePosInCIPBuffer_Detergent
    RoundedRectangle (75,174 35x20), "CIP5"
        tap fb.bTakePosInCIPBuffer_Full
    Lamp1 (6,38 29x28), variable: fb.bError, style: Lamp-Lamp1-Red
END_VISUALIZATION

// ---- 03 Project/10 Element/vis_FB_Element_CIP.TcVIS
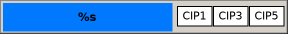
VISUALIZATION vis_FB_Element_CIP  // 288x34
VAR_IN_OUT
	fb: FB_Element;
END_VAR
    Rectangle (0,0 288x34)
    Textfield (2,2 171x30), "%s", text variable: fb.sElementID
    RoundedRectangle (177,6 35x20), "CIP1"
        tap fb.bTakePosInCIPBuffer_Partial
    RoundedRectangle (213,6 35x20), "CIP3"
        tap fb.bTakePosInCIPBuffer_Detergent
    RoundedRectangle (249,6 35x20), "CIP5"
        tap fb.bTakePosInCIPBuffer_Full
END_VISUALIZATION

// ---- 03 Project/11 Tank/vis_FB_ProductionTank.TcVIS
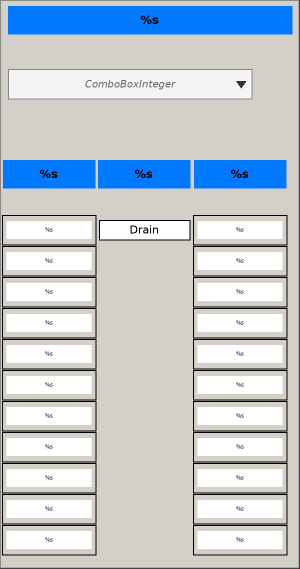
VISUALIZATION vis_FB_ProductionTank  // 300x569
VAR_IN_OUT
	fb: FB_ProductionTank;
END_VAR
    Rectangle (0,0 300x569)
    Textfield (7,5 286x30), "%s", text variable: fb.refElement.sElementID
    RoundedRectangle (99,220 91x20), "Drain"
        OnMouseClick: execute { fb.eReq:=E_Request_List.eDrain; }
    ComboBoxInteger (8,69 244x30), variable: fb.refElement.eState_Long, input disabled if: fb.refElement.bStateUpdate_Limited, text list: 'TextList_StateLong'
    Textfield (97,159 94x30), "%s", text variable: fb.eReq
    Textfield (193,159 94x30), "%s", text variable: fb.eProcess
    Textfield (2,159 94x30), "%s", text variable: fb.refElement.eState_Long, text list: 'TextList_StateLong', text index: fb.refElement.eState_Long
    Frame (2,215 94x30)
        shows vis_IconState(value := fb.refElement.eState_Long, reqValue := E_Element_State_Long.eStandby, text := 'Standby')
    Frame (2,246 94x30)
        shows vis_IconState(value := fb.refElement.eState_Long, reqValue := E_Element_State_Long.eNotClean, text := 'Not Clean')
    Frame (2,277 94x30)
        shows vis_IconState(value := fb.refElement.eState_Long, reqValue := E_Element_State_Long.eCIP_1_Rinzed, text := 'CIP1 Rinzed')
    Frame (2,308 94x30)
        shows vis_IconState(value := fb.refElement.eState_Long, reqValue := E_Element_State_Long.eCIP_2_Deterged, text := 'CIP2 Deterged')
    Frame (2,339 94x30)
        shows vis_IconState(value := fb.refElement.eState_Long, reqValue := E_Element_State_Long.eCIP_3_Deterged_Clean, text := 'CIP3 Deterged +')
    Frame (2,370 94x30)
        shows vis_IconState(value := fb.refElement.eState_Long, reqValue := E_Element_State_Long.eCIP_4_Sanitized, text := 'DisInfected')
    Frame (2,401 94x30)
        shows vis_IconState(value := fb.refElement.eState_Long, reqValue := E_Element_State_Long.eCIP_5_Done, text := 'CIP5 Done')
    Frame (2,432 94x30)
        shows vis_IconState(value := fb.refElement.eState_Long, reqValue := E_Element_State_Long.eWaterReady, text := 'WaterReady')
    Frame (2,463 94x30)
        shows vis_IconState(value := fb.refElement.eState_Long, reqValue := E_Element_State_Long.eReady, text := 'Ready')
    Frame (2,494 94x30)
        shows vis_IconState(value := fb.refElement.eState_Long, reqValue := E_Element_State_Long.eProduction, text := 'Production')
    Frame (2,525 94x30)
        shows vis_IconState(value := fb.refElement.eState_Long, reqValue := E_Element_State_Long.eExpired, text := 'Expired')
    Frame (193,215 94x30)
        shows vis_IconState(value := fb.eProcess, reqValue := E_Element_Process.eDrain, text := 'Draining')
    Frame (193,246 94x30)
        shows vis_IconState(value := fb.eProcess, reqValue := E_Element_Process.eWash_Recycle, text := 'Wash Recycle')
    Frame (193,277 94x30)
        shows vis_IconState(value := fb.eProcess, reqValue := E_Element_Process.eWash_Detergent, text := 'Wash Detergent')
    Frame (193,308 94x30)
        shows vis_IconState(value := fb.eProcess, reqValue := E_Element_Process.eWash_Water_1, text := 'Water 1')
    Frame (193,339 94x30)
        shows vis_IconState(value := fb.eProcess, reqValue := E_Element_Process.eWash_Sani, text := 'Wash DisInfection')
    Frame (193,370 94x30)
        shows vis_IconState(value := fb.eProcess, reqValue := E_Element_Process.eWash_Water_2, text := 'Water')
    Frame (193,401 94x30)
        shows vis_IconState(value := fb.eProcess, reqValue := E_Element_Process.eFill_Water, text := 'Filling Water')
    Frame (193,432 94x30)
        shows vis_IconState(value := fb.eProcess, reqValue := E_Element_Process.eDissolving, text := 'Dissolving')
    Frame (193,463 94x30)
        shows vis_IconState(value := fb.eProcess, reqValue := E_Element_Process.eConnectionToLine, text := 'Conn To Line')
    Frame (193,494 94x30)
        shows vis_IconState(value := fb.eProcess, reqValue := E_Element_Process.eDisconnection, text := 'Wash Detergent')
    Frame (193,525 94x30)
        shows vis_IconState(value := fb.eProcess, reqValue := E_Element_Process.eDrain, text := ' ')
END_VISUALIZATION

// ---- 03 Project/11 Tank/vis_IconState.TcVIS
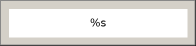
VISUALIZATION vis_IconState  // 196x46
VAR_IN_OUT
	value: INT;
END_VAR
VAR_INPUT
	reqValue: INT;
	text: STRING;	
END_VAR
    Rectangle (0,0 196x46), colour toggle: value=reqValue
    Textfield (8,8 180x30), "%s", text variable: text
        OnMouseClick: execute { value:=reqValue; }
END_VISUALIZATION

// ---- 03 Project/13 Weight control/TriBlender/VISUs/Main.TcVIS
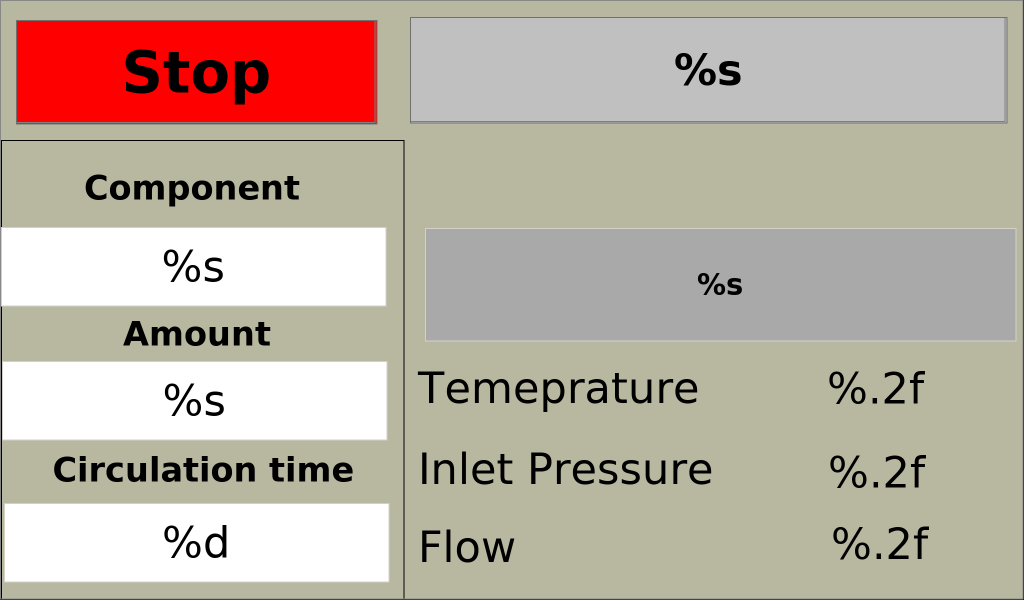
VISUALIZATION Main  // 1024x600
    Rectangle (0,0 1024x600)
    Button (16,20 361x104), "Stop"
    Button (410,17 597x106), "%s", text variable: prg_TriBlender.sStateDescription, input disabled if: prg_TriBlender.bDisableButton
        p2175578022: prg_TriBlender.wButtonColor
        OnMouseClick: execute { prg_TriBlender.bContinue:=TRUE; }
    Rectangle (1,140 403x460)
    Textfield (9,144 378x87), "Component", invisible if: prg_TriBlender.bDisableName
    Textfield (1,227 385x79), "%s", text variable: prg_TriBlender.stTriblender.sComponenetName, invisible if: prg_TriBlender.bDisableName
    Textfield (2,361 385x79), "%s", text variable: prg_TriBlender.stTriblender.sComponenetAmount, invisible if: prg_TriBlender.bDisableAmount
    Textfield (4,302 386x63), "Amount", invisible if: prg_TriBlender.bDisableAmount
    Textfield (7,441 393x57), "Circulation time", invisible if: prg_TriBlender.bDisableTime
    Textfield (4,503 385x79), "%d", text variable: prg_TriBlender.iCirculationTimeLeft, invisible if: prg_TriBlender.bDisableTime
    Textfield (425,228 591x113), "%s", text variable: prg_TriBlender.sStateInstructions
    Textfield (415,444 354x50), "Inlet Pressure"
    Textfield (765,441 223x63), "%.2f", text variable: prg_TriBlender.stTriblender.rPressure
    Textfield (415,522 354x50), "Flow"
    Textfield (767,517 225x54), "%.2f", text variable: prg_TriBlender.stTriblender.rFlow
    Textfield (415,363 354x50), "Temeprature"
    Textfield (764,365 223x47), "%.2f", text variable: prg_TriBlender.stTriblender.rTemp
END_VISUALIZATION

// ---- 03 Project/13 Weight control/TriBlender/VISUs/StartVisu.TcVIS
